// Simulation de toute la machine (docs/04 § 6.3)
{attribute 'qualified_only'}
VAR_GLOBAL
    bAllSimulated : BOOL;
    nSeed : UDINT := 16#2545F491;      // générateur pseudo-aléatoire des objets simulés (F_SimRandom)
END_VAR

(* stored: Version 1.1.0.1, ProductVersion 3.1.4024.12
   GVL GVL_Sim: Id {7faabaa4-fdef-5978-90b0-7d2b027d8c91} *)
